(* IEC 61131-3 sources: StewartPlatform/Class/VaranManager (part 4) *)

    if (ud_LenObjName + ud_LenStr) < VARAN_MUTEX_NAME_MAX_LENGTH then
      _strcat(dest:=#str_CombinedName[0], src:=#str_ObjName[0]);
    else
      _strncpy(dest:=#str_ObjNamePart1[0], src:= #str_ObjName[0], max:= VARAN_MUTEX_NAME_MAX_LENGTH - ud_LenStr - ud_SepLenStr - VARAN_MUTEX_NAME_END_LENGTH - 1);    // Copy Beginning of str_ObjName
      _strncpy(dest:=#str_ObjNamePart2[0], src:= #str_ObjName[ud_LenObjName-VARAN_MUTEX_NAME_END_LENGTH-1], max:=VARAN_MUTEX_NAME_END_LENGTH);  // Copy Last MUTEX_NAME_END_LENGTH Char of str_ObjName

      // Put the Mutex String together
      _strcat(dest:=#str_CombinedName[0], src:= #str_ObjNamePart1[0]);
      _strcat(dest:=#str_CombinedName[0], src:= VARAN_STR_MUTEX_NAME_SEPERATOR);
      _strcat(dest:=#str_CombinedName[0], src:= #str_ObjNamePart2[0]);
    end_if;

    pv_RetMutex := OS_MT_CreateSemaphore(MTSEMATYPE_MUTEX, 1, 0, #str_CombinedName[0]);

    if pv_RetMutex = nil then

      // If Create Mutex failed: Insert the this pointer into the string
      ud_LenCombObjName := _strlen(#str_CombinedName[0]);

      str_this[0] := '%';
      str_this[1] := 'm';
      _itoa(udNumber:=pthis$UDINT, pString:=#str_this[2]);
      ud_LenThis  := _strlen(src:=#str_this[0]);

      _strcpy(dest:=#str_CombinedName[ud_LenCombObjName-ud_LenThis], src:=#str_this[0]);

      pv_RetMutex := OS_MT_CreateSemaphore(MTSEMATYPE_MUTEX, 1, 0, #str_CombinedName[0]);

    end_if;

  end_if;

END_FUNCTION

FUNCTION GLOBAL VaranManager::MutexStart
  VAR_INPUT
    pMutex 	: pVoid;
  END_VAR

  if(pMutex <> NIL) then
    OS_MT_WAIT(pMutex);
  end_if;

END_FUNCTION

FUNCTION GLOBAL VaranManager::MutexStop
  VAR_INPUT
    pMutex 	: pVoid;
  END_VAR

  if(pMutex <> NIL) then
    OS_MT_SIGNAL(pMutex);
  end_if;

END_FUNCTION
#endif

FUNCTION VIRTUAL GLOBAL VaranManager::Control::NewInst
  VAR_INPUT
    pPara 	: ^CmdStruct;
    pResult 	: ^Results;
  END_VAR
  VAR_OUTPUT
    ret_code 	: IprStates;
  END_VAR
  VAR
    p_paraAddDO           : ^t_VM_CMD_AddDO;
    p_paraMovDO           : ^t_VM_CMD_AddMovDo;
    p_paraGetPointers     : ^t_VM_CMD_GetDataPointers;
    p_paraGetModuleHandel : ^t_VM_CMD_GetModuleHandle;
    PostInitRetcode       : iprStates;
    pHelpPostInit         : ^t_s_PostInitList;
    i                     : UINT;

    pHelp                 : ^void;  // This pointer to call newinst
    // local variables for the Requested HWTString
    pStr_HWTRequested     : ^CHAR;
    ui_HWTRequestedLength : UINT;
    us_HWTRequestedCurrIndex  : USINT;
    i_Req                 :UINT;
    // local variables for HWTStrings in the VM
    pStr_HWTVM            : ^CHAR;
    us_HWTVMLength        : USINT;
    i_VM                  : USINT;
    ud_ModuleIndex        : UDINT;
    b_ModuleFound         : BOOL;

    // local variables to safe currently found module
    pStr_HWTVMCurrent     : ^CHAR;
    ud_ModuleIndexCurrent : UDINT;

    TempArray         : ARRAY [0..SERNO_STRING_SIZE-1] OF USINT;
    a_HelpArray       : ARRAY[0..99] OF CHAR;
	  ud_StrSize : UDINT;
    ud_MaxStrSize : UDINT;
    sSPIIDHeader  : t_s_SPIListHeader;

    //local variables for dummy mux callback
    sd_retval           :DINT;
  END_VAR

  ret_code := READY;  // Overwritten on error

  CASE pPara^.uiCmd OF
//**********************************************************************************************************************************************************
    CMD_POST_INIT_CALL: // call from hwcontrol
      // Check Loader Version if function is supported
      if ops.uiLoaderVersion$UINT >= VM_POST_INIT_AVAILABLE then
        bPostInitActive := TRUE;

#ifdef _LSL_TARGETARCH_ARM  // IO Image only needed for ARM  CPUs
#ifdef VARAN_iSetOutputImage
        // the image is not copied from the shadow ram to the VM DPRAM so far => copy it
        if (b_IOImageWritten = FALSE) & b_IOImage then
          VARAN_iSetOutputImage(VaranManagerNr, VARAN_DOL_ASY);
          b_IOImageWritten := TRUE;
        end_if;
#endif
#endif

        // we wait here until the initialisation of the Varan Rt and the SDIAS Clients has been finished
        CyWork(0);

        if bPostInitModulesReady then
          ret_code := READY;
          bPostInitActive := FALSE;
        else
          ret_code := BUSY;
        end_if;
      else
        // Should be impossible as we never request a Postinit if the Loader version is incorrect.
        TRACE("(VaranManager::Control::NewInst) CMD_POST_INIT_CALL not supported with current Loader. Loader Version >= 02.02.137 is required");
        ret_code := ERROR;
      end_if;

//**********************************************************************************************************************************************************
    CMD_POST_INIT_RT_SYNC:
      // check if all modules are ready
      if WaitForSyncSendObjectsCnt then
        CyWork(0);

        ret_code := BUSY;
      end_if;

//**********************************************************************************************************************************************************
    CMD_POST_INIT_RT_READY:
      // check post init modules
      if PostInitModuleCnt then
        pHelpPostInit := #aPostInitList[0];
        for i := 0 to PostInitModuleCnt - 1 do

          //call class, if it's still not ready
          if pHelpPostInit^.p_This then
            PostInitRetcode := pHelpPostInit^.p_This^.NewInst(pPara, pResult);

            // only overwrite the ready returncode if the returncode from the post init objects is different to it
            if PostInitRetcode <> READY then
              ret_code := PostInitRetcode;
            end_if;
          end_if;

          // set pointer on next this pointer
          pHelpPostInit += sizeof(t_s_PostInitList);
        end_for;
      end_if;

      // if manager is disabled => return error
      if ManagerOn = 0 then
        ret_code := ERROR;

      // if we're not ready, return busy
      elsif us_RtStep <> _RtWork then
        ret_code := BUSY;

      elsif ret_code = READY then
        // everything ready
        b_PostInitRtSyncReady := TRUE;
      end_if;

//**********************************************************************************************************************************************************
    CMD_FORCE_POST_INIT_END:  // call from hwcontrol
      // HWControl has run into timeout and has ended the Post Init Phase
      // This call informs the VM thats the Phase has ended.
      bPostInitActive := FALSE;

//**********************************************************************************************************************************************************
    CMD_POST_INIT_DO_SORT:    // call from hwcontrol
      // sort safety DOs if there is more than 1
      if pPriorityList & pPriorityList^.pNext &
        b_PayloadSupport = false then     // OS Handles Priorities of DO if b_PayloadSupport = true

        SortCmdsByPriority();

#ifdef _LSL_TARGETARCH_ARM  // IO Image only needed for ARM  CPUs
#ifdef VARAN_iSetOutputImage
        // Varandata has to be written once after sorting the DOs
        if b_IOImage then
          VARAN_iSetOutputImage(VaranManagerNr, VARAN_DOL_ISO);
        end_if;
      else
        // Varandata has to be written once after adding the DOs even without sorting anything because we need the shadow RAM image in the VM DPRAM)
        if b_IOImage then
          VARAN_iSetOutputImage(VaranManagerNr, VARAN_DOL_ISO);
        end_if;
#endif
#endif
      end_if;
//**********************************************************************************************************************************************************
    CMD_GET_HARDWARE_TREE_ENTRY:

      pHelp                 := nil;  // This pointer to call newinst
      // local variables for the Requested HWTString
      ui_HWTRequestedLength := 0;
      us_HWTRequestedCurrIndex  := 0;
      i_Req                 := 0;
      // local variables for HWTStrings in the VM
      pStr_HWTVM            := NIL;
      us_HWTVMLength        := 0;
      i_VM                  := 0;
      ud_ModuleIndex        := 0;
      b_ModuleFound         := FALSE;

      // local variables to safe currently found module
      pStr_HWTVMCurrent     := NIL;
      ud_ModuleIndexCurrent := 0;

      ret_code := ERROR;
      pResult^.aData[0]$t_HWCGetHardwareTreeEntryOut.retcode := _HWC_RETVAL_ERROR_VARAN_MODULE_NOT_FOUND;

      pStr_HWTRequested     := pPara^.aPara[0]$t_HWCGetHardwareDiagnosisIn.pStr_HardewareTreeEntry;

      //First HWT Path
      if pStr_HWTRequested = nil then

        ud_VaranPosition := VM_OBJECT_PATH;

        // Return String of the Varanmanger
        ret_code := READY;
        pResult^.aData$t_HWCGetHardwareTreeEntryOut.retcode := _HWC_RETVAL_OK_HWTSTR_RETURNED;
        pResult^.aData[0]$t_HWCGetHardwareTreeEntryOut.pStr_NextHardewareTreeEntry := (#ud_VaranPosition)$^CHAR;

      // Only possible for VM own HWT Path
      elsif (pStr_HWTRequested^$USINT = 2) then

        if pStr_HWTRequested^$UDINT = VM_OBJECT_PATH then

          if s_ModuleList.p_ModuleList^ then
            // Return first Module in list
            ret_code := s_ModuleList.p_ModuleList^$p_VaranBase^.NewInst(pPara,pResult);
          else
            // VM was found but there are no modules connected
            ret_code := READY;
            pResult^.aData[0]$t_HWCGetHardwareTreeEntryOut.retcode := _HWC_RETVAL_OK_MODULE_FOUND;
          end_if;
        end_if;

      else

        //Search for module
        ui_HWTRequestedLength     := (pStr_HWTRequested)$^UINT^ + 1;  //+1 because we compare the strings, 2 byte length
        us_HWTRequestedCurrIndex  := pPara^.aPara[0]$t_HWCGetHardwareDiagnosisIn.us_current_index;

        ud_ModuleIndex := 0;
        b_ModuleFound := FALSE;

        //loop over all modules
        while (ud_ModuleIndex < s_ModuleList.ud_NrOfModules) &
              (b_ModuleFound = FALSE) do

          pStr_HWTVM := (s_ModuleList.p_PositionList+ (ud_ModuleIndex * 4))^$^CHAR;  // 4 = SizeOf(^CHAR)

          if pStr_HWTVM  then
            us_HWTVMLength := pStr_HWTVM^;  //First byte is length

            i_Req := us_HWTRequestedCurrIndex;
            i_Vm  := 1;

            //Loop over strings
            while i_Req <= ui_HWTRequestedLength &
                  i_Vm  <= us_HWTVMLength do

              if (pStr_HWTRequested + i_Req)^ <> (pStr_HWTVM + i_Vm)^ then // Compare byte
                // Strings are not equal
                exit;
              end_if;

              i_Req += 1;
              i_VM  += 1;
            end_while;

            if (i_Req <= ui_HWTRequestedLength ) &                        // End of requested string was not reached
               (i_Vm = us_HWTVMLength + 1) &                              // And end of compared string reached
               ( (pStr_HWTRequested + i_Req)^ and HWT_ESCAPE_SEQU ) then  // Escape sequece found in Requested string

              b_ModuleFound := TRUE;

//              pPara^.aPara[0]$t_HWCGetHardwareDiagnosisIn.us_current_index   := i_Req$USINT;
//              pPara^.aPara[0]$t_HWCGetHardwareDiagnosisIn.us_current_length  := (ui_HWTRequestedLength - i_Req)$USINT;
              exit;
            end_if;

            if (i_Vm = us_HWTVMLength + 1) & (i_Req = ui_HWTRequestedLength + 1) then   // All Bytes and Length are equal
              b_ModuleFound := TRUE;
#ifdef HWK_SHOW_PRAGMA_MESSAGES
              #pragma message("LanSte 26.06.2014 16:11 \ check")
#endif

//              pPara^.aPara[0]$t_HWCGetHardwareDiagnosisIn.us_current_index  := i_Req$USINT - 1;  // -1 because we increased over max length at the end of the while loop
//              pPara^.aPara[0]$t_HWCGetHardwareDiagnosisIn.us_current_length := 1; // Last entry of string was reached, index points to last entry
              exit;
            end_if;

          end_if;

          ud_ModuleIndex += 1;  // Select next Module

        end_while;

        if b_ModuleFound then

          // Call module again incase it is an extension module
          pHelp := s_ModuleList.p_ModuleList + sizeof(p_VaranBase) * ud_ModuleIndex;
          ret_code := pHelp^$p_VaranBase^.NewInst(pPara,pResult);

          // Return if new HWT String was found
          if ret_code = READY &
             pResult^.aData[0]$t_HWCGetHardwareDiagnosisOut.retcode = _HWC_RETVAL_OK_HWTSTR_RETURNED then
            return;
          end_if;

          ud_ModuleIndex += 1;  // Select next Module
          ud_ModuleIndexCurrent := ud_ModuleIndex;

          b_ModuleFound := TRUE;  // Only set to enter loop

          while (ud_ModuleIndexCurrent < s_ModuleList.ud_NrOfModules) &
                (b_ModuleFound = TRUE) do

            pStr_HWTVMCurrent := (s_ModuleList.p_PositionList+ (ud_ModuleIndexCurrent * 4))^$^CHAR ;  // 4 = SizeOf(^CHAR)

            if pStr_HWTVMCurrent then

              // Check if module has already been called (multiple entries in list)
              ud_ModuleIndex := 0;
              b_ModuleFound := FALSE;

              //loop over all modules to search for duplicates
              while (ud_ModuleIndex < ud_ModuleIndexCurrent &
                     b_ModuleFound = FALSE) do

                pStr_HWTVM := (s_ModuleList.p_PositionList+ (ud_ModuleIndex * 4))^$^CHAR ;  // 4 = SizeOf(^CHAR)

                if pStr_HWTVM then

                  // Compare string length
                  if pStr_HWTVMCurrent^ = pStr_HWTVM^ then

                    // Compare string content
                    if _memcmp( ptr1 := pStr_HWTVMCurrent + 1,
                                ptr2 := pStr_HWTVM +1,
                                cntr := pStr_HWTVMCurrent^) = 0 then

                      // Multiple entry, Check next Module
                      b_ModuleFound := TRUE;
                      ud_ModuleIndexCurrent += 1;
                      exit;

                    end_if;
                  end_if;
                end_if;

                ud_ModuleIndex += 1;

              end_while;

              if b_ModuleFound = FALSE then
                exit; // Non duplicate entry
              end_if;

            else  // if pStr_HWTVMCurrent then
              ud_ModuleIndexCurrent += 1;
            end_if;

          end_while;

          if b_ModuleFound = FALSE then
            // Call Class
            pHelp := s_ModuleList.p_ModuleList + sizeof(p_VaranBase) * ud_ModuleIndexCurrent;
            ret_code := pHelp^$p_VaranBase^.NewInst(pPara,pResult);
          end_if;

        else
          pResult^.aData[0]$t_HWCGetHardwareDiagnosisOut.retcode := _HWC_RETVAL_ERROR_VARAN_MODULE_NOT_FOUND;
          ret_code := ERROR;
        end_if;

      end_if;

//**********************************************************************************************************************************************************
    CMD_GET_HARDWARE_DIAGNOSIS:

      pHelp                 := nil;  // This pointer to call newinst
      // local variables for the Requested HWTString
      ui_HWTRequestedLength := 0;
      us_HWTRequestedCurrIndex  := 0;
      i_Req                 := 0;
      // local variables for HWTStrings in the VM
      pStr_HWTVM            := NIL;
      us_HWTVMLength        := 0;
      i_VM                  := 0;
      ud_ModuleIndex        := 0;
      b_ModuleFound         := FALSE;

      ret_code := ERROR;
      pResult^.aData[0]$t_HWCGetHardwareDiagnosisOut.retcode := _HWC_RETVAL_ERROR;

      pStr_HWTRequested     := pPara^.aPara[0]$t_HWCGetHardwareDiagnosisIn.pStr_HardewareTreeEntry;

      if pStr_HWTRequested then

        // Check for VM String
        if (pStr_HWTRequested)$^UINT^ = 2 then

          if (pStr_HWTRequested)$^UDINT^ = VM_OBJECT_PATH then

            TempArray[0] := 0;

            if this <> p_this then
              //Reset statemachine
              eSPISSW := _GetVendorName;
              //Save This pointer
              p_this := this;

              // Reset Flags
              bDiagnosisDataAvailableFlags.HWVersion   := FALSE;
              bDiagnosisDataAvailableFlags.VendorName  := FALSE;
              bDiagnosisDataAvailableFlags.DeviceName  := FALSE;
              bDiagnosisDataAvailableFlags.OrderingNo  := FALSE;
              bDiagnosisDataAvailableFlags.LicenseNo   := FALSE;
              bDiagnosisDataAvailableFlags.SerialNo    := FALSE;
            end_if;

            case eSPISSW of
            	_GetVendorName:
                ret_code$DINT := GetSPIDataFromID(  p_us_position_info:=#TempArray[0]
                                                  , udListID:= VM_SPI_VENDOR_NAME_ID
                                                  , pData:= #a_VendorName[0]
                                                  , udRequDataLength:= sizeof(a_VendorName)
                                                  , pIDHeader:= #sSPIIDHeader
                                                  );

                if ret_code = READY then

                  // Null Termination ----------------------------------------
                  ud_StrSize    := sSPIIDHeader.ListLength;
                  ud_MaxStrSize := sizeof(a_VendorName);

                  pResult^.aData[0]$t_HWCGetHardwareDiagnosisOut.pStr_VendorName  := (#a_VendorName)$^CHAR; // Will be overwritten if this pointer is not equal

                  (pResult^.aData[0]$t_HWCGetHardwareDiagnosisOut.pStr_VendorName + ud_MaxStrSize)^ := 0;
                  if ud_StrSize < ud_MaxStrSize then
                    (pResult^.aData[0]$t_HWCGetHardwareDiagnosisOut.pStr_VendorName + ud_StrSize)^ := 0;
                  end_if;

                  bDiagnosisDataAvailableFlags.VendorName := TRUE;

                  eSPISSW := _GetSerialNo;
                  ret_code := BUSY;
                else
                  pResult^.aData[0]$t_HWCGetHardwareDiagnosisOut.retcode := _HWC_RETVAL_ERROR_VARAN_SPI_ACCESS_FAILED;
                  //set SSW to SPI Data Ready, because we return the values which are already in the HWK
                  eSPISSW := _SPIDataReady;
                  ret_code := BUSY;
                end_if;

              _GetSerialNo:
                ret_code$DINT := GetSPIDataFromID(  p_us_position_info:=#TempArray[0]
                                                  , udListID:= VM_SPI_SERIALNO_ID
                                                  , pData:= #a_SerialNo[0]
                                                  , udRequDataLength:= sizeof(a_SerialNo)
                                                  , pIDHeader:= #sSPIIDHeader
                                                  );

                if ret_code = READY then

                  // Null Termination ----------------------------------------
                  ud_StrSize    := sSPIIDHeader.ListLength;
                  ud_MaxStrSize := sizeof(a_SerialNo);

                  pResult^.aData[0]$t_HWCGetHardwareDiagnosisOut.pStr_SerialNo  := (#a_SerialNo)$^CHAR; // Will be overwritten if this pointer is not equal

                  (pResult^.aData[0]$t_HWCGetHardwareDiagnosisOut.pStr_SerialNo + ud_MaxStrSize)^ := 0;
                  if ud_StrSize < ud_MaxStrSize then
                    (pResult^.aData[0]$t_HWCGetHardwareDiagnosisOut.pStr_SerialNo + ud_StrSize)^ := 0;
                  end_if;

                  bDiagnosisDataAvailableFlags.SerialNo := TRUE;

                  eSPISSW := _GetDeviceName;
                  ret_code := BUSY;
                else
                  pResult^.aData[0]$t_HWCGetHardwareDiagnosisOut.retcode := _HWC_RETVAL_ERROR_VARAN_SPI_ACCESS_FAILED;
                  //set SSW to SPI Data Ready, because we return the values which are already in the HWK
                  eSPISSW := _SPIDataReady;
                  ret_code := BUSY;
                end_if;

            	_GetDeviceName:
                ret_code$DINT := GetSPIDataFromID(  p_us_position_info:=#TempArray[0]
                                                  , udListID:= VM_SPI_DEVICE_NAME_ID
                                                  , pData:= #a_DeviceName[0]
                                                  , udRequDataLength:= sizeof(a_DeviceName)
                                                  , pIDHeader:= #sSPIIDHeader
                                                  );

                if ret_code = READY then

                  // Null Termination ----------------------------------------
                  ud_StrSize    := sSPIIDHeader.ListLength;
                  ud_MaxStrSize := sizeof(a_DeviceName);

                  pResult^.aData[0]$t_HWCGetHardwareDiagnosisOut.pStr_DeviceName  := (#a_DeviceName)$^CHAR; // Will be overwritten if this pointer is not equal

                  (pResult^.aData[0]$t_HWCGetHardwareDiagnosisOut.pStr_DeviceName + ud_MaxStrSize)^ := 0;
                  if ud_StrSize < ud_MaxStrSize then
                    (pResult^.aData[0]$t_HWCGetHardwareDiagnosisOut.pStr_DeviceName + ud_StrSize)^ := 0;
                  end_if;

                  bDiagnosisDataAvailableFlags.DeviceName := TRUE;

                  eSPISSW := _GetOrderingNo;
                  ret_code := BUSY;
                else
                  pResult^.aData[0]$t_HWCGetHardwareDiagnosisOut.retcode := _HWC_RETVAL_ERROR_VARAN_SPI_ACCESS_FAILED;
                  //set SSW to SPI Data Ready, because we return the values which are already in the HWK
                  eSPISSW := _SPIDataReady;
                  ret_code := BUSY;
                end_if;

            	_GetOrderingNo:
                ret_code$DINT := GetSPIDataFromID(  p_us_position_info:=#TempArray[0]
                                                  , udListID:= VM_SPI_ORDERING_NO_ID
                                                  , pData:= #a_OrderingNo[0]
                                                  , udRequDataLength:= sizeof(a_OrderingNo)
                                                  , pIDHeader:= #sSPIIDHeader
                                                  );

                if ret_code = READY then

                  // Null Termination ----------------------------------------
                  ud_StrSize    := sSPIIDHeader.ListLength;
                  ud_MaxStrSize := sizeof(a_OrderingNo);

                  pResult^.aData[0]$t_HWCGetHardwareDiagnosisOut.pStr_OrderingNo  := (#a_OrderingNo)$^CHAR; // Will be overwritten if this pointer is not equal

                  (pResult^.aData[0]$t_HWCGetHardwareDiagnosisOut.pStr_OrderingNo + ud_MaxStrSize)^ := 0;
                  if ud_StrSize < ud_MaxStrSize then
                    (pResult^.aData[0]$t_HWCGetHardwareDiagnosisOut.pStr_OrderingNo + ud_StrSize)^ := 0;
                  end_if;

                  bDiagnosisDataAvailableFlags.OrderingNo := TRUE;

                  eSPISSW := _GetLicenseNoHWVersion;
                  ret_code := BUSY;
                else
                  pResult^.aData[0]$t_HWCGetHardwareDiagnosisOut.retcode := _HWC_RETVAL_ERROR_VARAN_SPI_ACCESS_FAILED;
                  //set SSW to SPI Data Ready, because we return the values which are already in the HWK
                  eSPISSW := _SPIDataReady;
                  ret_code := BUSY;
                end_if;

            	_GetLicenseNoHWVersion:

                ret_code$DINT := GetSPIDataFromID(  p_us_position_info:=#TempArray[0]
                                                  , udListID:= VM_SPI_IDENTIFICATION_LIST
                                                  , pData:= #a_HelpArray[0]
                                                  , udRequDataLength:= sizeof(udHWVersion) + sizeof(udLicenseNo)
                                                  , pIDHeader:= #sSPIIDHeader
                                                  , udOffset := 8
                                                  );

                udLicenseNo := a_HelpArray[0]$UDINT;
                udHWVersion := a_HelpArray[4]$UDINT;

                if ret_code = READY then
                  bDiagnosisDataAvailableFlags.LicenseNo := TRUE;
                  bDiagnosisDataAvailableFlags.HWVersion := TRUE;
                  eSPISSW := _SPIDataReady;
                  ret_code := BUSY;
                else
                  pResult^.aData[0]$t_HWCGetHardwareDiagnosisOut.retcode := _HWC_RETVAL_ERROR_VARAN_SPI_ACCESS_FAILED;
                  //set SSW to SPI Data Ready, because we return the values which are already in the HWK
                  eSPISSW := _SPIDataReady;
                  ret_code := BUSY;
                end_if;

            	_SPIDataReady:
                //Don't reset statemachine because if we have the same this pointer we don't have to make spi Accesses again
                //eSPISSW := _GetVendorName;

                //Data which is already in HWK available
                if p_NodeInfo then

                  pResult^.aData$t_HWCGetHardwareDiagnosisOut.hd_FPGAVersion  := to_udint(p_NodeInfo^.ucFPGAVersion);
                  pResult^.aData$t_HWCGetHardwareDiagnosisOut.ud_DeviceID     := to_udint(p_NodeInfo^.uiDeviceID);
                  pResult^.aData$t_HWCGetHardwareDiagnosisOut.ud_VendorID     := to_udint(p_NodeInfo^.uiVendorID);
                end_if;

                if bDiagnosisDataAvailableFlags.VendorName then
                  pResult^.aData[0]$t_HWCGetHardwareDiagnosisOut.pStr_VendorName  := (#a_VendorName)$^CHAR;
                end_if;

                if bDiagnosisDataAvailableFlags.HWVersion & bDiagnosisDataAvailableFlags.LicenseNo then
                  pResult^.aData[0]$t_HWCGetHardwareDiagnosisOut.hd_HWVersion     := udHWVersion;
                  pResult^.aData[0]$t_HWCGetHardwareDiagnosisOut.ud_LicenseNo      := udLicenseNo;
                end_if;

                if bDiagnosisDataAvailableFlags.DeviceName then
                  pResult^.aData[0]$t_HWCGetHardwareDiagnosisOut.pStr_DeviceName  := (#a_DeviceName)$^CHAR;
                end_if;

                if bDiagnosisDataAvailableFlags.OrderingNo then
                  pResult^.aData[0]$t_HWCGetHardwareDiagnosisOut.pStr_OrderingNo  := (#a_OrderingNo)$^CHAR;
                end_if;

                if bDiagnosisDataAvailableFlags.SerialNo then
                  pResult^.aData[0]$t_HWCGetHardwareDiagnosisOut.pStr_SerialNo := (#a_SerialNo)$^CHAR;
                end_if;

                ret_code := READY;
                pResult^.aData[0]$t_HWCGetHardwareDiagnosisOut.retcode := _HWC_RETVAL_OK;

            end_case;
          end_if;

          return;
        end_if;

        ui_HWTRequestedLength     := (pStr_HWTRequested)$^UINT^ + 1;  //+1 because we compare the strings, 2 byte length
        us_HWTRequestedCurrIndex  := pPara^.aPara[0]$t_HWCGetHardwareDiagnosisIn.us_current_index;

        ud_ModuleIndex := 0;
        b_ModuleFound := FALSE;

        //loop over all modules
        while (ud_ModuleIndex < s_ModuleList.ud_NrOfModules) &
              (b_ModuleFound = FALSE) do

          pStr_HWTVM := (s_ModuleList.p_PositionList+ (ud_ModuleIndex * 4))^$^CHAR ;  // 4 = SizeOf(^CHAR)

          if pStr_HWTVM  then
            us_HWTVMLength := pStr_HWTVM^;  //First byte is length

            i_Req := us_HWTRequestedCurrIndex;
            i_Vm  := 1;

            //Loop over strings
            while i_Req <= ui_HWTRequestedLength &
                  i_Vm  <= us_HWTVMLength do

//              if (pStr_HWTRequested + i_Req)^ and HWT_ESCAPE_SEQU then  // Check for Escape Sequenze
//                b_ModuleFound := TRUE;
//                exit;
//              end_if;

              if (pStr_HWTRequested + i_Req)^ <> (pStr_HWTVM + i_Vm)^ then // Compare byte
                // Strings are not equal
                exit;
              end_if;

              i_Req += 1;
              i_VM  += 1;
            end_while;

//            #pragma message("LanSte 18.06.2014 18:23 \ Index Update testen")
//            if b_ModuleFound then // Escape Sequence was found
//
//              pPara^.aPara[0]$t_HWCGetHardwareDiagnosisIn.us_current_index   := i_Req$USINT;
//              pPara^.aPara[0]$t_HWCGetHardwareDiagnosisIn.us_current_length  := (ui_HWTRequestedLength - i_Req)$USINT;
//              exit;
//
//            end_if;

            if (i_Req <= ui_HWTRequestedLength ) &                        // End of requested string was not reached
            (i_Vm = us_HWTVMLength + 1) &                                 // And end of compared string reached
               ( (pStr_HWTRequested + i_Req)^ and HWT_ESCAPE_SEQU ) then  // Escape sequece found in Requested string

              b_ModuleFound := TRUE;
              pPara^.aPara[0]$t_HWCGetHardwareDiagnosisIn.us_current_index   := i_Req$USINT;
              pPara^.aPara[0]$t_HWCGetHardwareDiagnosisIn.us_current_length  := (ui_HWTRequestedLength - i_Req)$USINT;
              exit;
            end_if;

            if (i_Vm = us_HWTVMLength + 1) & (i_Req = ui_HWTRequestedLength + 1) then   // All Bytes and Length are equal
              b_ModuleFound := TRUE;
              pPara^.aPara[0]$t_HWCGetHardwareDiagnosisIn.us_current_index  := i_Req$USINT - 1;  // -1 because we increased over max length at the end of the while loop
              pPara^.aPara[0]$t_HWCGetHardwareDiagnosisIn.us_current_length := 1; // Last entry of string was reached, index points to last entry
              exit;
            end_if;

          end_if;

          ud_ModuleIndex += 1;  // Select next Module

        end_while;

        if b_ModuleFound then
          // Call Class
          pHelp := s_ModuleList.p_ModuleList + sizeof(p_VaranBase) * ud_ModuleIndex;
          ret_code := pHelp^$p_VaranBase^.NewInst(pPara,pResult);
        else
          pResult^.aData[0]$t_HWCGetHardwareDiagnosisOut.retcode := _HWC_RETVAL_ERROR_VARAN_MODULE_NOT_FOUND;
          ret_code := ERROR;
        end_if;

      end_if;

//**********************************************************************************************************************************************************
    VM_CMD_NEED_POST_INIT_CALL: // call from varan client
      // Check Loader Version if function is supported
      if ops.uiLoaderVersion$UINT >= VM_POST_INIT_AVAILABLE then

        // store this pointer of the module
        aPostInitList[PostInitModuleCnt].p_This := pPara^.aPara[0]$p_VaranBase;

        // remember if we have to wait for DOs to be created
        aPostInitList[PostInitModuleCnt].Settings := pPara^.aPara[1]$BSINT;
        if aPostInitList[PostInitModuleCnt].Settings.Wait4DOCreation then
          WaitForPostInitObjectsCnt += 1;
          if aPostInitList[PostInitModuleCnt].Settings.Wait4MoveDOCreation then
            WaitForPostInitMoveObjectsCnt += 1;
          end_if;
        end_if;

        // remember if we have to wait for the sync of this module
        if aPostInitList[PostInitModuleCnt].Settings.Wait4SyncSend then
          WaitForSyncSendObjectsCnt += 1;
        end_if;

        aPostInitList[PostInitModuleCnt].b_CallMe := TRUE;

        // return index for this module
        pResult^.uiLng := 2;
        pResult^.aData[0]$UINT := PostInitModuleCnt;

        // increase number of post init modules
        PostInitModuleCnt += 1;

        // we're no longer ready with post init. we have to wait until all modules from the list are finished
        bPostInitModulesReady := FALSE;
      else
        TRACE("(VaranManager::Control::NewInst) VM_CMD_NEED_POST_INIT_CALL not supported with current Loader. Loader Version >= 02.02.137 is required");
        ret_code := ERROR;
      end_if;

//**********************************************************************************************************************************************************
    VM_CMD_POST_INIT_FINISHED: // call from varan client
      // Check Loader Version if function is supported
      if ops.uiLoaderVersion$UINT >= VM_POST_INIT_AVAILABLE then

        // only relevant during last Init
        if PostInitModuleCnt then
          // check if it's a valid index
          if pPara^.aPara[1]$UINT < VM_MAX_POST_INIT_MODULES then
            // check if our local this pointer matches this object
            if pPara^.aPara[0]$p_VaranBase = aPostInitList[pPara^.aPara[1]$UINT].p_This then
              // increase number of ready objects
              PostInitModuleReadyCnt += 1;
//              aPostInitList[pPara^.aPara[1]$UINT].b_CallMe := FALSE;

              // check if it's an object we were waiting for
              if aPostInitList[pPara^.aPara[1]$UINT].Settings.Wait4DOCreation then
                aPostInitList[pPara^.aPara[1]$UINT].Settings.Wait4DOCreation := FALSE;

                if WaitForPostInitObjectsCnt then
                  WaitForPostInitObjectsCnt -= 1;
                else
                  TRACE("(VaranManager::Control::NewInst) There is already no more post init object to wait for! (VM_CMD_POST_INIT_FINISHED)");
                  ret_code := ERROR;
                end_if;
              end_if;

              // check if it's an object we were waiting for
              if aPostInitList[pPara^.aPara[1]$UINT].Settings.Wait4MoveDOCreation then
                aPostInitList[pPara^.aPara[1]$UINT].Settings.Wait4MoveDOCreation := FALSE;

                if WaitForPostInitMoveObjectsCnt then
                  WaitForPostInitMoveObjectsCnt -= 1;
                else
                  TRACE("(VaranManager::Control::NewInst) There is already no more post init object to wait for (create move DOs)! (VM_CMD_POST_INIT_FINISHED)");
                  ret_code := ERROR;
                end_if;
              end_if;

              // on last init we check if all modules which need to have finished their init
              if PostInitModuleReadyCnt = PostInitModuleCnt then
                bPostInitModulesReady := TRUE;
              end_if;
            else
              TRACE("(VaranManager::Control::NewInst) This pointer of post init module given doesn't match locally stored this pointer for this index!");
              ret_code := ERROR;
            end_if;
          else
            TRACE("(VaranManager::Control::NewInst) Invalid index of post init module given!");
            ret_code := ERROR;
          end_if;
        else
          TRACE("(VaranManager::Control::NewInst) More modules ready with last init than expected");
          ret_code := ERROR;
        end_if;
      else
        TRACE("(VaranManager::Control::NewInst) VM_CMD_POST_INIT_FINISHED not supported with current Loader. Loader Version >= 02.02.137 is required");
        ret_code := ERROR;
      end_if;

//**********************************************************************************************************************************************************
    VM_CMD_IS_PAYLOAD_SUPPORTED:  // to get the status of PayloadSupport
      pResult^.aData[0]$BOOL := b_PayloadSupport;

//**********************************************************************************************************************************************************
    VM_CMD_DO_CREATION_FINISHED: // a post-init module is finished with creating DOs
      // Check Loader Version if function is supported
      if ops.uiLoaderVersion$UINT >= VM_POST_INIT_AVAILABLE then

        // only relevant during last Init
        if PostInitModuleCnt then
          // check if it's a valid index
          if pPara^.aPara[1]$UINT < VM_MAX_POST_INIT_MODULES then
            // check if our local this pointer matches this object
            if pPara^.aPara[0]$p_VaranBase = aPostInitList[pPara^.aPara[1]$UINT].p_This then
              // check if it's an object we were waiting for
              if aPostInitList[pPara^.aPara[1]$UINT].Settings.Wait4DOCreation then
                aPostInitList[pPara^.aPara[1]$UINT].Settings.Wait4DOCreation := FALSE;

                if WaitForPostInitObjectsCnt then
                  WaitForPostInitObjectsCnt -= 1;
                else
                  TRACE("(VaranManager::Control::NewInst) There is already no more post init object to wait for!");
                  ret_code := ERROR;
                end_if;
              else
                TRACE("(VaranManager::Control::NewInst) Module finished with DO creation, where  There is already no more post init object to wait for!");
                ret_code := ERROR;
              end_if;
            else
              TRACE("(VaranManager::Control::NewInst) This pointer of post init module given doesn't match locally stored this pointer for this index!");
              ret_code := ERROR;
            end_if;
          else
            TRACE("(VaranManager::Control::NewInst) Invalid index of post init module given!");
            ret_code := ERROR;
          end_if;
        else
          TRACE("(VaranManager::Control::NewInst) More modules ready with last init than expected");
          ret_code := ERROR;
        end_if;
      else
        TRACE("(VaranManager::Control::NewInst) VM_CMD_DO_CREATION_FINISHED not supported with current Loader. Loader Version >= 02.02.137 is required");
        ret_code := ERROR;
      end_if;

//**********************************************************************************************************************************************************
    VM_CMD_MOVE_DO_CREATION_FINISHED:
      // Check Loader Version if function is supported
      if ops.uiLoaderVersion$UINT >= VM_POST_INIT_AVAILABLE then

        // only relevant during last Init
        if PostInitModuleCnt then
          // check if it's a valid index
          if pPara^.aPara[1]$UINT < VM_MAX_POST_INIT_MODULES then
            // check if our local this pointer matches this object
            if pPara^.aPara[0]$p_VaranBase = aPostInitList[pPara^.aPara[1]$UINT].p_This then
              // check if it's an object we were waiting for
              if aPostInitList[pPara^.aPara[1]$UINT].Settings.Wait4MoveDOCreation then
                aPostInitList[pPara^.aPara[1]$UINT].Settings.Wait4MoveDOCreation := FALSE;

                if WaitForPostInitMoveObjectsCnt then
                  WaitForPostInitMoveObjectsCnt -= 1;
                else
                  TRACE("(VaranManager::Control::NewInst) There is already no more post init object to wait for (create move DOs)!");
                  ret_code := ERROR;
                end_if;
              else
                TRACE("(VaranManager::Control::NewInst) Module finished with move DO creation, where  There is already no more post init object to wait for!");
                ret_code := ERROR;
              end_if;
            else
              TRACE("(VaranManager::Control::NewInst) This pointer of post init module given doesn't match locally stored this pointer for this index! (Move DOs)");
              ret_code := ERROR;
            end_if;
          else
            TRACE("(VaranManager::Control::NewInst) Invalid index of post init module given! (Move DOs)");
            ret_code := ERROR;
          end_if;
        else
          TRACE("(VaranManager::Control::NewInst) More modules ready with last init than expected (Move DOs)");
          ret_code := ERROR;
        end_if;
      else
        TRACE("(VaranManager::Control::NewInst) VM_CMD_MOVE_DO_CREATION_FINISHED not supported with current Loader. Loader Version >= 02.02.137 is required (Move DOs)");
        ret_code := ERROR;
      end_if;

//**********************************************************************************************************************************************************
    VM_CMD_DO_MEM_READY: // check if all post init objects are finished with creating DOs
      // if we're not in post init or the varan manager has finished waiting for post init objects => the DO memory is ready
      if WaitForPostInitObjectsCnt = 0 then
        pResult^.aData[4] := TRUE;
      else
        pResult^.aData[4] := FALSE;
      end_if;

//**********************************************************************************************************************************************************
    VM_CMD_MOVE_DO_MEM_READY: // check if all post init objects are finished with creating move DOs
      // if we're not in post init or the varan manager has finished waiting for post init objects => the move DO memory is ready
      if WaitForPostInitMoveObjectsCnt = 0 then
        pResult^.aData[4] := TRUE;
      else
        pResult^.aData[4] := FALSE;
      end_if;

//**********************************************************************************************************************************************************
    VM_CMD_SYNC_SEND_READY:
      // only work on it if the post init rt hasn't been finished, otherwise we would have the log messages if modules are plugged at runtime
      if b_PostInitRtSyncReady = FALSE then
        // Check Loader Version if function is supported
        if ops.uiLoaderVersion$UINT >= VM_POST_INIT_AVAILABLE then
          // only relevant during last Init
          if PostInitModuleCnt then
            // check if it's a valid index
            if pPara^.aPara[1]$UINT < VM_MAX_POST_INIT_MODULES then
              // check if our local this pointer matches this object
              if pPara^.aPara[0]$p_VaranBase = aPostInitList[pPara^.aPara[1]$UINT].p_This then
                // check if it's an object we were waiting for
                if aPostInitList[pPara^.aPara[1]$UINT].Settings.Wait4SyncSend then
                  aPostInitList[pPara^.aPara[1]$UINT].Settings.Wait4SyncSend := FALSE;

                  if WaitForSyncSendObjectsCnt then
                    WaitForSyncSendObjectsCnt -= 1;
                  else
                    TRACE("(VaranManager::Control::NewInst) There is already no more post init object to wait for (sync send ready)!");
                    ret_code := ERROR;
                  end_if;
                else
                  TRACE("(VaranManager::Control::NewInst) Module finished with sync send ready, where  There is already no more post init object to wait for!");
                  ret_code := ERROR;
                end_if;
              else
                TRACE("(VaranManager::Control::NewInst) This pointer of post init module given doesn't match locally stored this pointer for this index! (Move DOs)");
                ret_code := ERROR;
              end_if;
            else
              TRACE("(VaranManager::Control::NewInst) Invalid index of post init module given! (sync send ready)");
              ret_code := ERROR;
            end_if;
          else
            TRACE("(VaranManager::Control::NewInst) More modules ready with last init than expected (sync send ready)");
            ret_code := ERROR;
          end_if;
        else
          TRACE("(VaranManager::Control::NewInst) VM_CMD_MOVE_DO_CREATION_FINISHED not supported with current Loader. Loader Version >= 02.02.137 is required (Move DOs)");
          ret_code := ERROR;
        end_if;
      end_if;

//**********************************************************************************************************************************************************
    VM_CMD_SET_MUX_THIS: // ignore this command, it's only for the VaranMux classes
      ret_code := ERROR; // return error => command not handled

//**********************************************************************************************************************************************************
    VM_CMD_INSTALL_DUMMY_CALLBACK:

      if pPara^.aPara[0] >= 4 * sizeof(DINT) then

        sd_retval := AddObjectCallback(p_us_position_info:=pPara^.aPara[1]$^USINT
                        , ud_action_ptr:= pPara^.aPara[2]$UDINT
                        , ud_thisp:= pPara^.aPara[3]$UDINT
                        , sd_required:= pPara^.aPara[4]);
      else

        TRACE("(VaranManager::Control::NewInst) VM_CMD_INSTALL_DUMMY_CALLBACK. Length of NewInst Commando is invalid");
      end_if;

//**********************************************************************************************************************************************************
    else    // Commands for Payload
      if b_PayloadSupport then

        pResult^.uiLng := sizeof(DINT);
        pResult^.aData[0]$DINT := VM_CMD_NOT_IMPLEMENTED; // Default Return code, must be overwritten by induvidual methods

        CASE pPara^.uiCmd OF

        //*****************************************************************************
          VM_CMD_GET_MODULE_HANDLE :
            p_paraGetModuleHandel := (pPara^.aPara[0])$^t_VM_CMD_GetModuleHandle;

            pResult^.aData[0]$DINT := GetModuleHandle(  p_us_PositionInfo := p_paraGetModuleHandel^.p_us_position_info
                                                      , p_ud_ModuleHandle := p_paraGetModuleHandel^.p_ud_module_handle);

        //*****************************************************************************
          VM_CMD_ADD_DO :
            p_paraAddDO := (pPara^.aPara[0])$^t_VM_CMD_AddDO;
            pResult^.aData[0]$DINT := AddPayloadDO( p_ud_DoHandle                 := p_paraAddDO^.p_ud_DoHandle
                                                  , ud_NodeHandle                 := p_paraAddDO^.ud_ModuleHandle
                                                  , ud_DoRequired                 := p_paraAddDO^.ud_b_DoRequired
                                                  , ud_DolType                    := p_paraAddDO^.ud_DolType
                                                  , ud_Command                    := p_paraAddDO^.ud_Command
                                                  , ud_Priority                   := p_paraAddDO^.ud_Priority
                                                  , ud_PrescalerCounterThreshold  := p_paraAddDO^.ud_PreScalerCounterThreshold
                                                  , ud_PrescalerCounterStartValue := p_paraAddDO^.ud_PreScalerCounterStartValue
                                                  , ud_ReadOffset                 := p_paraAddDO^.ud_OffsetRead
                                                  , ud_ReadLength                 := p_paraAddDO^.ud_LengthRead
                                                  , ud_WriteOffset                := p_paraAddDO^.ud_OffsetWrite
                                                  , ud_WriteLength                := p_paraAddDO^.ud_LengthWrite
                                                  , ud_Filter                     := p_paraAddDO^.ud_Filter
                                                  , ud_Slices                     := p_paraAddDO^.ud_Slices
                                                  , ud_WritePayloadType           := p_paraAddDO^.ud_WritePayloadType);

        //*****************************************************************************
          VM_CMD_ADD_MOV_DO :
            p_paraMovDO := (pPara^.aPara[0])$^t_VM_CMD_AddMovDo;
            pResult^.aData[0]$DINT := AddPayloadMoveDO( p_ud_DoHandle                 := p_paraMovDO^.p_ud_DoHandle
                                                      , ud_bDoRequired                := p_paraMovDO^.ud_b_DoRequired
                                                      , ud_DolType                    := p_paraMovDO^.ud_DolType
                                                      , ud_Priority                   := p_paraMovDO^.ud_Priority
                                                      , ud_PrescalerCounterThreshold  := p_paraMovDO^.ud_PreScalerCounterThreshold
                                                      , ud_PrescalerCounterStartValue := p_paraMovDO^.ud_PreScalerCounterStartValue
                                                      , ud_hSourceReadDoHandle        := p_paraMovDO^.ud_SourceReadDoHandle
                                                      , ud_ReadOffset                 := p_paraMovDO^.ud_SourceReadOffset
                                                      , ud_hDestinationWriteDoHandle  := p_paraMovDO^.ud_DestinationWriteDoHandle
                                                      , ud_WriteOffset                := p_paraMovDO^.ud_DestinationWriteOffset
                                                      , ud_MoveDataLength             := p_paraMovDO^.ud_LengthMove);

        //*****************************************************************************
          VM_CMD_GET_DATA_POINTERS  :
            p_paraGetPointers := (pPara^.aPara[0])$^t_VM_CMD_GetDataPointers;
            pResult^.aData[0]$DINT := GetDataPointers(  ud_hDoHandle  := p_paraGetPointers^.ud_DoHandle
                                                      , pp_ReadData   := p_paraGetPointers^.p_ud_ReadData$^pVoid
                                                      , pp_WriteData  := p_paraGetPointers^.p_ud_WriteData$^pVoid);

        //*****************************************************************************
          VM_CMD_IS_DMA_ACTIVE :
            if PayloadFrame then
              pResult^.aData[0]$BOOL := TRUE;
            else
              pResult^.aData[0]$BOOL := FALSE;
            end_if;

          else
            ret_code := ERROR;
        END_CASE;

      else
        pResult^.uiLng := sizeof(DINT);
        pResult^.aData[0]$DINT := VM_CMD_NOT_IMPLEMENTED;
        TRACE("(VaranManager::Control::NewInst) Unknown command!");
        ret_code := ERROR;
      end_if;

  END_CASE;

END_FUNCTION

FUNCTION VaranManager::TurnOffIsoTask
  VAR
    s_PropertyValuePair : LSL_PROPERTY_VALUE_PAIR;
  END_VAR

  if b_PayloadSupport &
     _RTOSVersion >= VM_FULL_PAYLOAD_AVAILABLE  then
    s_PropertyValuePair.udPropertyId    := VM_PROP_TASK_STATE_ISO;
    s_PropertyValuePair.udPropertyValue := TK_STATE_STOPPED;
    MULTI_VARAN_iSetNodeProperties( hNodeHandle           := vmNodeHandle
                                  , udPropertyCount       := 1
                                  , psPropertyValuePairs  := #s_PropertyValuePair);
  else
    p_ManagerStructure^.ucTCEnable := p_ManagerStructure^.ucTCEnable AND VM_DISABLE_ISO_TASK;
  end_if;

END_FUNCTION

FUNCTION VaranManager::AddPayloadDO
  VAR_INPUT
    p_ud_DoHandle 	: ^UDINT;
    ud_NodeHandle 	: UDINT;
    ud_DoRequired 	: UDINT;
    ud_DolType 	: UDINT;
    ud_Command 	: UDINT;
    ud_Priority 	: UDINT;
    ud_PrescalerCounterThreshold 	: UDINT;
    ud_PrescalerCounterStartValue 	: UDINT;
    ud_ReadOffset 	: UDINT;
    ud_ReadLength 	: UDINT;
    ud_WriteOffset 	: UDINT;
    ud_WriteLength 	: UDINT;
    ud_Filter 	: UDINT;
    ud_Slices 	: UDINT;
    ud_WritePayloadType :  UDINT;
  END_VAR
  VAR_OUTPUT
    sd_retval 	: DINT;
  END_VAR
  VAR
    TempMem             :  UDINT;
    TempMemWr           :  UDINT;
  END_VAR

#ifdef VM_DEBUG_PAYLOAD
  if b_PayloadSupport = false then
    // This method is not suppored without payload
    ((0)$^USINT)^ := 0;
  end_if;
#endif

  //look if we Manager is on
  if ( ManagerOn ) then
    //look if we must execute Cyclic DOL list
    if ( ud_DolType = VARAN_DOL_ASY ) then
      s_CyHandles.b_ExecuteDOL := TRUE;			//set flag to execut Dol list
    end_if;

    sd_retval := MULTI_VARAN_iAddDo(  phDoHandle    := p_ud_DoHandle
                                    , hNodeHandle   := ud_NodeHandle
                                    , bDoRequired   := ud_DoRequired
                                    , udDolType     := ud_DolType
                                    , udCommand     := ud_Command
                                    , udPriority    := ud_Priority
                                    , udPrescalerCounterThreshold   := ud_PrescalerCounterThreshold
                                    , udPrescalerCounterStartValue  := ud_PrescalerCounterStartValue
                                    , udReadOffset  := ud_ReadOffset
                                    , udReadLength  := ud_ReadLength
                                    , udWriteOffset := ud_WriteOffset
                                    , udWriteLength := ud_WriteLength
                                    , udFilter      := ud_Filter
                                    , udSlices      := ud_Slices
                                    , udWritePayloadType := ud_WritePayloadType$LSL_WRITE_PAYLOAD_TYPE);

    //look if an error occured
    if ( sd_retval <> VARANMANAGER_OK ) then
      s_ErrorVaranManager.f_AddRdDO := SetVaranDOError( sd_Error 		:= sd_retval
                                                      , b_manager_off	:= TRUE
                                                      , b_log			:= TRUE
                                                      );
    else

      if PayloadFrame then  // Use PayloadFrame because, b_PayloadSupport only shows the interface used.
                            // Payload DO Mem Calculaition +++++++++++++++++++++++++++++++++++++++++++++++++++++++++++++++++++++++++++++++++++++++++++++++++++++++++++++++++++++++++++++++++++++++++
        case ud_Command of

            VARAN_CMD_CONTROL_READ,
            VARAN_CMD_MEMORY_READ:      // Read DO -------------------------------------------------------------------------------------------------------------------------------
                // 1 Byte Status + n Byte (Load data read) + 0 to 3 Byte (compensate missalignment)
                TempMem := 1 + ud_ReadLength;

                // 1 Byte Control
                TempMemWr := 1;

                // Increase for variable DO
                if ud_WritePayloadType > WR_PLD_TYPE_STANDARD$UDINT then
                  TempMemWr += 16#0D;
                end_if;

                case ud_DolType of
                // **************************************************
                  VARAN_DOL_DA:
                    DPRAM_Used.DA_Rd          += TempMem + TempMemWr + SIZE_PAYLOAD_FRAME_HEADER_DO;
                    DPRAM_Used_Payload.DA_Rd  += TempMem;
                    DPRAM_Used_Payload.DA_Wr  += TempMemWr;
                    DOCounter.DA_Rd  += 1;

                // **************************************************
                  VARAN_DOL_ISO:
                    DPRAM_Used.ISO_Rd         += TempMem + TempMemWr + SIZE_PAYLOAD_FRAME_HEADER_DO;
                    DPRAM_Used_Payload.ISO_Rd += TempMem;
                    DPRAM_Used_Payload.ISO_Wr += TempMemWr;
                    DOCounter.ISO_Rd  += 1;

                // **************************************************
                  VARAN_DOL_ASY:
                    DPRAM_Used.ASY_Rd         += TempMem + TempMemWr + SIZE_PAYLOAD_FRAME_HEADER_DO;
                    DPRAM_Used_Payload.ASY_Rd += TempMem;
                    DPRAM_Used_Payload.ASY_Wr += TempMemWr;
                    DOCounter.ASY_Rd  += 1;

                // **************************************************
                  VARAN_DOL_ADMIN:
                    DPRAM_Used.Admin_Rd         += TempMem + TempMemWr + SIZE_PAYLOAD_FRAME_HEADER_DO;
                    DPRAM_Used_Payload.Admin_Rd += TempMem;
                    DPRAM_Used_Payload.ASY_Wr   += TempMemWr;
                    DOCounter.Admin_Rd += 1;

                // **************************************************
                  VARAN_DOL_IRQ:
                    DPRAM_Used.IRQ_Rd         += TempMem + TempMemWr + SIZE_PAYLOAD_IRQ_FRAME_HEADER_DO;
                    DPRAM_Used_Payload.IRQ_Rd += TempMem;
                    DPRAM_Used_Payload.IRQ_Wr += TempMemWr;
                    DOCounter.IRQ_Rd  += 1;
                end_case;

                DPRAM_Used_Payload.Payload_Read += TempMem;
                DPRAM_Used_Payload.Payload_Write += TempMemWr;

                if ud_DolType <> VARAN_DOL_IRQ then
                  DPRAM_Used.Total  += TempMem + TempMemWr + SIZE_PAYLOAD_FRAME_HEADER_DO;
                  DPRAM_Used_Payload.Payload_Header += SIZE_PAYLOAD_FRAME_HEADER_DO;
                else
                  DPRAM_Used.Total  += TempMem + TempMemWr + SIZE_PAYLOAD_IRQ_FRAME_HEADER_DO;
                  DPRAM_Used_Payload.Payload_Header += SIZE_PAYLOAD_IRQ_FRAME_HEADER_DO;
                end_if;

                DPRAM_Used_Payload.Total  += TempMem + TempMemWr;

                DOCounter.Total   += 1;

            VARAN_CMD_CONTROL_WRITE,
            VARAN_CMD_MEMORY_WRITE:     // Write DO -------------------------------------------------------------------------------------------------------------------------------
                // 1 Byte Control + n Byte (Load data read) + 0 to 3 Byte (compensate missalignment)
                TempMemWr := 1 + ud_WriteLength;

                // Increase for variable DO
                if ud_WritePayloadType > WR_PLD_TYPE_STANDARD$UDINT then
                  TempMemWr += 16#0D;
                end_if;

                // 1 Byte Status in Read DPRAM
                TempMem := 1;

                case ud_DolType of
                // **************************************************
                  VARAN_DOL_DA:
                    DPRAM_Used.DA_Wr            += TempMem + TempMemWr + SIZE_PAYLOAD_FRAME_HEADER_DO;
                    DPRAM_Used_Payload.DA_Rd    += TempMem;
                    DPRAM_Used_Payload.DA_Wr    += TempMemWr;
                    DOCounter.DA_Wr  += 1;

                // **************************************************
                  VARAN_DOL_ISO:
                    DPRAM_Used.ISO_Wr           += TempMem + TempMemWr + SIZE_PAYLOAD_FRAME_HEADER_DO;
                    DPRAM_Used_Payload.ISO_Rd   += TempMem;
                    DPRAM_Used_Payload.ISO_Wr   += TempMemWr;
                    DOCounter.ISO_Wr += 1;

                // **************************************************
                  VARAN_DOL_ASY:
                    DPRAM_Used.ASY_Wr           += TempMem + TempMemWr + SIZE_PAYLOAD_FRAME_HEADER_DO;
                    DPRAM_Used_Payload.ASY_Rd   += TempMem;
                    DPRAM_Used_Payload.ASY_Wr   += TempMemWr;
                    DOCounter.ASY_Wr  += 1;

                // **************************************************
                  VARAN_DOL_ADMIN:
                    DPRAM_Used.Admin_Wr         += TempMem + TempMemWr + SIZE_PAYLOAD_FRAME_HEADER_DO;
                    DPRAM_Used_Payload.Admin_Rd += TempMem;
                    DPRAM_Used_Payload.Admin_Wr += TempMemWr;
                    DOCounter.Admin_Wr  += 1;

                // **************************************************
                  VARAN_DOL_IRQ:
                    DPRAM_Used.IRQ_Wr           += TempMem + TempMemWr + SIZE_PAYLOAD_IRQ_FRAME_HEADER_DO;
                    DPRAM_Used_Payload.ISO_Rd   += TempMem;
                    DPRAM_Used_Payload.IRQ_Wr   += TempMemWr;
                    DOCounter.IRQ_Wr  += 1;

                end_case;

                DPRAM_Used_Payload.Payload_Read += TempMem;
                DPRAM_Used_Payload.Payload_Write += TempMemWr;

                if ud_DolType <> VARAN_DOL_IRQ then
                  DPRAM_Used.Total  += TempMem + TempMemWr + SIZE_PAYLOAD_FRAME_HEADER_DO;
                  DPRAM_Used_Payload.Payload_Header += SIZE_PAYLOAD_FRAME_HEADER_DO;
                else
                  DPRAM_Used.Total  += TempMem + TempMemWr + SIZE_PAYLOAD_IRQ_FRAME_HEADER_DO;
                  DPRAM_Used_Payload.Payload_Header += SIZE_PAYLOAD_IRQ_FRAME_HEADER_DO;
                end_if;

                DPRAM_Used_Payload.Total  += TempMem + TempMemWr;
                DOCounter.Total   += 1;

            VARAN_CMD_CONTROL_READ_WRITE,
            VARAN_CMD_MEMORY_READ_WRITE:// Read/Write DO -------------------------------------------------------------------------------------------------------------------------------
                // 1 Byte Control + n Byte (Load data read) + 0 to 3 Byte (compensate missalignment) x2
                TempMem := 1 + ud_ReadLength;

                TempMemWr := 1 + ud_WriteLength;

                // Increase for variable DO
                if ud_WritePayloadType = WR_PLD_TYPE_RW_ACCESS_CONFIGURABLE$UDINT then
                  TempMemWr += 16#13;
                elsif ud_WritePayloadType > WR_PLD_TYPE_STANDARD$UDINT then
                  TempMemWr += 16#0D;
                end_if;

                case ud_DolType of
                // **************************************************
                  VARAN_DOL_DA:
                    DPRAM_Used.DA_RdWr += TempMem + TempMemWr + SIZE_PAYLOAD_FRAME_HEADER_DO;
                    DPRAM_Used_Payload.DA_Rd += TempMem;
                    DPRAM_Used_Payload.DA_Wr += TempMemWr;
                    DOCounter.DA_RdWr  += 1;

                // **************************************************
                  VARAN_DOL_ISO:
                    DPRAM_Used.ISO_RdWr += TempMem + TempMemWr + SIZE_PAYLOAD_FRAME_HEADER_DO;
                    DPRAM_Used_Payload.ISO_Rd += TempMem;
                    DPRAM_Used_Payload.ISO_Wr += TempMemWr;

                    DOCounter.ISO_RdWr  += 1;

                // **************************************************
                  VARAN_DOL_ASY:
                    DPRAM_Used.ASY_RdWr += TempMem + TempMemWr + SIZE_PAYLOAD_FRAME_HEADER_DO;
                    DPRAM_Used_Payload.ASY_Rd += TempMem;
                    DPRAM_Used_Payload.ASY_Wr += TempMemWr;
                    DOCounter.ASY_RdWr  += 1;

                // **************************************************
                  VARAN_DOL_ADMIN:
                    DPRAM_Used.Admin_RdWr += TempMem + TempMemWr + SIZE_PAYLOAD_FRAME_HEADER_DO;
                    DPRAM_Used_Payload.Admin_Rd += TempMem;
                    DPRAM_Used_Payload.Admin_Wr += TempMemWr;
                    DOCounter.Admin_RdWr  += 1;

                // **************************************************
                  VARAN_DOL_IRQ:
                    DPRAM_Used.IRQ_RdWr += TempMem + TempMemWr + SIZE_PAYLOAD_IRQ_FRAME_HEADER_DO;
                    DPRAM_Used_Payload.IRQ_Rd += TempMem;
                    DPRAM_Used_Payload.IRQ_Wr += TempMemWr;
                    DOCounter.IRQ_RdWr  += 1;

                end_case;

                DPRAM_Used_Payload.Payload_Read += TempMem;
                DPRAM_Used_Payload.Payload_Write += TempMemWr;

                if ud_DolType <> VARAN_DOL_IRQ then
                  DPRAM_Used.Total  += TempMem + TempMemWr + SIZE_PAYLOAD_FRAME_HEADER_DO;
                  DPRAM_Used_Payload.Payload_Header += SIZE_PAYLOAD_FRAME_HEADER_DO;
                else
                  DPRAM_Used.Total  += TempMem + TempMemWr + SIZE_PAYLOAD_IRQ_FRAME_HEADER_DO;
                  DPRAM_Used_Payload.Payload_Header += SIZE_PAYLOAD_IRQ_FRAME_HEADER_DO;
                end_if;

                DPRAM_Used_Payload.Total += TempMem + TempMemWr;
                DOCounter.Total   += 1;

        end_case;
      else    // Standard DO Mem Calculation +++++++++++++++++++++++++++++++++++++++++++++++++++++++++++++++++++++++++++++++++++++++++++++++++++++++++++++++++++++++++++++++++++++++++

        case ud_Command of

            VARAN_CMD_CONTROL_READ,
            VARAN_CMD_MEMORY_READ:      // Read DO -------------------------------------------------------------------------------------------------------------------------------
                // 32 Byte (Header) + 6 Byte (1 Byte Cmd, 4 Byte Addr, 1 Byte Len) + 1 Byte (Response) + n Byte (Load data read) + 0 to 3 Byte (compensate missalignment)
                TempMem := 32 + 6 + 1 + ud_ReadLength;
                if (TempMem MOD 4) then
                  TempMem := TempMem + (4 - (TempMem MOD 4)); //increase memory, up to a value, which could be divided by 4
                end_if;

                case ud_DolType of
                // **************************************************
                  VARAN_DOL_DA:
                                DPRAM_Used.DA_Rd += TempMem;
                                DOCounter.DA_Rd  += 1;
                // **************************************************
                  VARAN_DOL_ISO:
                                DPRAM_Used.ISO_Rd += TempMem;
                                DOCounter.ISO_Rd  += 1;
                // **************************************************
                  VARAN_DOL_ASY:
                                DPRAM_Used.ASY_Rd += TempMem;
                                DOCounter.ASY_Rd  += 1;
                // **************************************************
                  VARAN_DOL_ADMIN:
                                DPRAM_Used.Admin_Rd += TempMem;
                                DOCounter.Admin_Rd  += 1;
                // **************************************************
                  VARAN_DOL_IRQ:
                                DPRAM_Used.IRQ_Rd += TempMem;
                                DOCounter.IRQ_Rd  += 1;
                end_case;

                DPRAM_Used.Total  += TempMem;
                DOCounter.Total   += 1;

            VARAN_CMD_CONTROL_WRITE,
            VARAN_CMD_MEMORY_WRITE:     // Write DO -------------------------------------------------------------------------------------------------------------------------------
                //32 Byte (Header) + 6 Byte (1 Byte Cmd, 4 Byte Addr, 1 Byte Len) + 1 Byte (Response) + n Byte (load data write) + 0 to 3 Byte (compensate missalignment)
                  TempMem := 32 + 6 + 1 + ud_WriteLength;
                  if (TempMem MOD 4) then
                    TempMem := TempMem + (4 - (TempMem MOD 4)); //increase memory, up to a value, which could be divided by 4
                  end_if;

                  case ud_DolType of
                  // **************************************************
                    VARAN_DOL_DA:
                                  DPRAM_Used.DA_Wr += TempMem;
                                  DOCounter.DA_Wr  += 1;
                  // **************************************************
                    VARAN_DOL_ISO:
                                  DPRAM_Used.ISO_Wr += TempMem;
                                  DOCounter.ISO_Wr  += 1;
                  // **************************************************
                    VARAN_DOL_ASY:
                                  DPRAM_Used.ASY_Wr += TempMem;
                                  DOCounter.ASY_Wr  += 1;
                  // **************************************************
                    VARAN_DOL_ADMIN:
                                  DPRAM_Used.Admin_Wr += TempMem;
                                  DOCounter.Admin_Wr  += 1;
                  // **************************************************
                    VARAN_DOL_IRQ:
                                  DPRAM_Used.IRQ_Wr += TempMem;
                                  DOCounter.IRQ_Wr  += 1;
                  end_case;

                  DPRAM_Used.Total  += TempMem;
                  DOCounter.Total   += 1;

            VARAN_CMD_CONTROL_READ_WRITE,
            VARAN_CMD_MEMORY_READ_WRITE:// Read/Write DO -------------------------------------------------------------------------------------------------------------------------------
                  //32 Byte (Header) + 11 Byte (1 Byte Cmd, 4 Byte RdAddr, 1 Byte RdLen, 4 Byte WrAddr, 1 Byte WrLen) + 1 Byte (Response) + n Byte (load data read) + n Byte (load data write) + 0 to 3 Byte (compensate missalignment)
                  TempMem := 32 + 11 + 1 + ud_ReadLength + ud_WriteLength;
                  if (TempMem MOD 4) then
                    TempMem := TempMem + (4 - (TempMem MOD 4)); //increase memory, up to a value, which could be divided by 4
                  end_if;

                  case ud_DolType of
                  // **************************************************
                    VARAN_DOL_DA:
                                  DPRAM_Used.DA_RdWr += TempMem;
                                  DOCounter.DA_RdWr  += 1;
                  // **************************************************
                    VARAN_DOL_ISO:
                                  DPRAM_Used.ISO_RdWr += TempMem;
                                  DOCounter.ISO_RdWr  += 1;
                  // **************************************************
                    VARAN_DOL_ASY:
                                  DPRAM_Used.ASY_RdWr += TempMem;
                                  DOCounter.ASY_RdWr  += 1;
                  // **************************************************
                    VARAN_DOL_ADMIN:
                                  DPRAM_Used.Admin_RdWr += TempMem;
                                  DOCounter.Admin_RdWr  += 1;
                  // **************************************************
                    VARAN_DOL_IRQ:
                                  DPRAM_Used.IRQ_RdWr += TempMem;
                                  DOCounter.IRQ_RdWr  += 1;
                  end_case;

                  DPRAM_Used.Total  += TempMem;
                  DOCounter.Total   += 1;

        end_case;

      end_if; // +++++++++++++++++++++++++++++++++++++++++++++++++++++++++++++++++++++++++++++++++++++++++++++++++++++++++++++++++++++++++++++++++++++++++++++++++++++++++++++++++++++++++++++++++

    end_if;
  else
    sd_retval := -100;	//Manager is off
  end_if;
END_FUNCTION

FUNCTION VaranManager::AddPayloadMoveDO
  VAR_INPUT
    p_ud_DoHandle 	: ^UDINT;
    ud_bDoRequired 	: UDINT;
    ud_DolType 	: UDINT;
    ud_Priority 	: UDINT;
    ud_PrescalerCounterThreshold 	: UDINT;
    ud_PrescalerCounterStartValue 	: UDINT;
    ud_hSourceReadDoHandle 	: UDINT;
    ud_ReadOffset 	: UDINT;
    ud_hDestinationWriteDoHandle 	: UDINT;
    ud_WriteOffset 	: UDINT;
    ud_MoveDataLength 	: UDINT;
  END_VAR
  VAR_OUTPUT
    sd_retval 	: DINT;
  END_VAR

#ifdef VM_DEBUG_PAYLOAD
  if b_PayloadSupport = false then
    // This method is not suppored without payload
    ((0)$^USINT)^ := 0;
  end_if;
#endif

  //look if we must execute Cyclic DOL list
  if ( ud_DolType = VARAN_DOL_ASY ) then
    s_CyHandles.b_ExecuteDOL := TRUE;			//set flag to execut Dol list
  end_if;

  sd_retval := MULTI_VARAN_iAddMoveDo(  phDoHandle                    := p_ud_DoHandle
                                      , bDoRequired                   := ud_bDoRequired
                                      , udDolType                     := ud_DolType
                                      , udPriority                    := ud_Priority
                                      , udPrescalerCounterThreshold   := ud_PrescalerCounterThreshold
                                      , udPrescalerCounterStartValue  := ud_PrescalerCounterStartValue
                                      , hSourceReadDoHandle           := ud_hSourceReadDoHandle
                                      , udReadOffset                  := ud_ReadOffset
                                      , hDestinationWriteDoHandle     := ud_hDestinationWriteDoHandle
                                      , udWriteOffset                 := ud_WriteOffset
                                      , udMoveDataLength              := ud_MoveDataLength);
  //look if an error occured
  if ( sd_retval <> VARANMANAGER_OK ) then
    s_ErrorVaranManager.f_AddRdDO := SetVaranDOError( sd_Error      := sd_retval
                                                    , b_manager_off := TRUE
                                                    , b_log         := TRUE
                                                    );
  else
    // Payload Move DO Mem Calculation
    if ( ud_DolType = VARAN_DOL_ASY ) then
      DPRAM_Used.ASY_Mov          += sizeof(LSL_VARANFRAMEPAYLOADMOVEHEADER);
      DPRAM_Used_Payload.ASY_Rd   += 1; // 1 Byte status
      DPRAM_Used_Payload.ASY_Wr   += sizeof(LSL_VARANFRAMEMOVEWRITEPAYLOAD);
      DOCounter.ASY_Mov           += 1;
    else
      DPRAM_Used.ISO_Mov          += sizeof(LSL_VARANFRAMEPAYLOADMOVEHEADER);
      DPRAM_Used_Payload.ISO_Rd   += 1; // 1 Byte status
      DPRAM_Used_Payload.ISO_Wr   += sizeof(LSL_VARANFRAMEMOVEWRITEPAYLOAD);
      DOCounter.ISO_Mov           += 1;
    end_if;

    DPRAM_Used.Total          += sizeof(LSL_VARANFRAMEPAYLOADMOVEHEADER) + 1 + sizeof(LSL_VARANFRAMEMOVEWRITEPAYLOAD);  // Header + Read Statusbyte + Write Payload
    DPRAM_Used_Payload.Total  += 1 + sizeof(LSL_VARANFRAMEMOVEWRITEPAYLOAD);  // Read Statusbyte + Write Payload
    DOCounter.Total           += 1;
  end_if;

END_FUNCTION

FUNCTION VaranManager::GetDataPointers
  VAR_INPUT
    ud_hDoHandle 	: UDINT;
    pp_ReadData 	: ^pVoid;
    pp_WriteData 	: ^pVoid;
  END_VAR
  VAR_OUTPUT
    sd_retval 	: DINT;
  END_VAR

#ifdef VM_DEBUG_PAYLOAD
  if b_PayloadSupport = false then
    // This method is not suppored without payload
    ((0)$^USINT)^ := 0;
  end_if;
#endif

  // if there is no VARAN Interface available, we would crash at the call
  if pMultiVaran = NIL then
    sd_retval := VARANMANAGER_DRIVER_NOT_EXISTS;
    return;
  end_if;

  sd_retval :=  MULTI_VARAN_iGetDataPointers( hDoHandle   := ud_hDoHandle
                                            , ppvReadData := pp_ReadData
                                            , ppvWriteData:= pp_WriteData);

END_FUNCTION

FUNCTION VaranManager::GetModuleHandle
  VAR_INPUT
    p_us_PositionInfo 	: ^USINT;
    p_ud_ModuleHandle 	: ^UDINT;
  END_VAR
  VAR_OUTPUT
    sd_retval 	: DINT;
  END_VAR

  // if there is no VARAN Interface available, we would crash at the call
  if pMultiVaran = NIL then
    sd_retval := VARANMANAGER_DRIVER_NOT_EXISTS;
    return;
  end_if;

  sd_retval := MULTI_VARAN_iGetNodeHandle(  udManagerNumber := VaranManagerNr
                                          , pszHardwarePath := p_us_PositionInfo
                                          , phNodeHandle    := p_ud_ModuleHandle);

END_FUNCTION

FUNCTION VaranManager::AddObjectCallback
	VAR_INPUT
		p_us_position_info 	: ^USINT;
		ud_action_ptr 	: UDINT;
		ud_thisp 	: UDINT;
		sd_required 	: DINT;
	END_VAR
	VAR_OUTPUT
		sd_retval 	: DINT;
	END_VAR
VAR
  ud_NodeHandle       :UDINT;
END_VAR

  if State = _NoVaranInterface then
    sd_retval := -100;
    return;
  end_if;
  //get right required flag
  if ( sd_required ) then
    sd_required := VARAN_DEVICE_REQUIRED;
  else
    sd_required := VARAN_DEVICE_DEFAULT;
  end_if;

    if b_PayloadSupport &
         _RTOSVersion >= VM_FULL_PAYLOAD_AVAILABLE  then
      sd_retval := MULTI_VARAN_iGetNodeHandle(  udManagerNumber := VaranManagerNr
                                              , pszHardwarePath := p_us_position_info
                                              , phNodeHandle    := #ud_NodeHandle);

      if sd_retval <> VARANMANAGER_OK then
        return;
      end_if;

      //call OS - function to set callback
      sd_retval := MULTI_VARAN_iSetApplicationCallback( hNodeHandle           := ud_NodeHandle
                                                      , pfApplicationCallback := ud_action_ptr$pvoid
                                                      , pvUserData            := ud_thisp$pvoid
                                                      , udRequired            := sd_required$UDINT);

    elsif pVaran then

      //call OS - function to set callback
      sd_retval := VARAN_iSetObjectCallback	( uiManager := VaranManagerNr
                                            , pucNode   := p_us_position_info
                                            , uiCallback:= ud_action_ptr
                                            , uiThis    := ud_thisp
                                            , uiRequired:= sd_required$UDINT
                                            );
    end_if;

  //look for an error
  if ( sd_retval <> VARANMANAGER_OK ) then
    s_ErrorVaranManager.f_SetObjectCallback := SetVaranDOError	( sd_Error 		:= sd_retval
                                                                , b_manager_off	:= TRUE
                                                                , b_log			:= TRUE
                                                                );
  end_if;

END_FUNCTION

FUNCTION VIRTUAL VaranManager::LogValue
	VAR_INPUT
		pString 	: ^CHAR;
		Value 	: UDINT;
		Value2 	: UDINT;(* := 16#FFFFFFFF *)
		Value3 	: UDINT;(* := 16#FFFFFFFF *)
	END_VAR
  VAR
    TempStr       : ARRAY [0..99] OF CHAR;
    TempStr2      : ARRAY [0..99] OF CHAR;
    TempStr3      : ARRAY [0..99] OF CHAR;
    TraceVal      : USINT;
    sz_name       : ARRAY [ 0..255 ] OF CHAR;
    TmpWithObjName: ARRAY [ 0..255 ] OF CHAR;
  END_VAR

  // number of values
  TraceVal := 1;

  _itoa(Value, #TempStr[0]);

  if pString <> NIL then
    _GetObjName( this, #sz_name[ 0 ] );
    _strcpy(dest:=#TmpWithObjName[0], src:="ObjectName ");
    _strcat(dest:=#TmpWithObjName[0], src:=#sz_name[0]);
    _strcat(dest:=#TmpWithObjName[0], src:=": ");
    _strcat(dest:=#TmpWithObjName[0], src:=pString);

    if Value2 <> 16#FFFFFFFF then
      _itoa(Value2, #TempStr2[0]);
      TraceVal += 1;
    end_if;

    if Value3 <> 16#FFFFFFFF then
      _itoa(Value3, #TempStr3[0]);
      TraceVal += 1;
    end_if;

    case TraceVal of
      1:MyTrace(pFormat:=#TmpWithObjName[0], pTxt0:=#TempStr[0], pTxt1:=NIL, pTxt2:=NIL);
      2:MyTrace(pFormat:=#TmpWithObjName[0], pTxt0:=#TempStr[0], pTxt1:=#TempStr2[0], pTxt2:=NIL);
      3:MyTrace(pFormat:=#TmpWithObjName[0], pTxt0:=#TempStr[0], pTxt1:=#TempStr2[0], pTxt2:=#TempStr3[0]);
    end_case;
  else
    MyTrace(pFormat:="<invalid string>", pTxt0:=NIL, pTxt1:=NIL, pTxt2:=NIL);
  end_if;

END_FUNCTION

FUNCTION VIRTUAL VaranManager::MyTrace
	VAR_INPUT
		pFormat 	: ^CHAR;
		pTxt0 	: ^CHAR;
		pTxt1 	: ^CHAR;
		pTxt2 	: ^CHAR;
	END_VAR
  VAR
    nLen      : UDINT;
    pChr      : ^CHAR;
    nTxt      : UDINT;
    nRpl      : UDINT;
    pTxt      : ^CHAR;
    pText     : ^CHAR;
    FormText  : ARRAY [0 .. 255] OF CHAR;
  END_VAR

  // this method is a workaround for the TRACE message limitation problem

  pText := #FormText[0];

  _memset(dest:=#FormText[0], usByte:=0, cntr:=256); // to keep the zero termination

  _strncpy(pText, pFormat, 250);
  nLen  := _strlen(pText);
  pChr  := pText;

  WHILE nLen DO
    IF pChr^ = '{' THEN         // works for the first 10 replacement texts (single digit numbers)
      nTxt  := (pChr+1)^ - '0';
      CASE nTxt OF
        0:  pTxt  := pTxt0;
        1:  pTxt  := pTxt1;
        2:  pTxt  := pTxt2;
      ELSE
        pTxt  := "INV";
      END_CASE;
      nRpl  := _strlen(pTxt);
      if nLen - 3 + nRpl > 250 then
        pTxt := "LEN";  // replace the replacement text with "LEN" to see that we're out of length for this string
        nRpl := 3;
      end_if;
      _memmove(pChr + nRpl, pChr + 3, nLen);
      _memcpy(pChr, pTxt, nRpl);
      pChr  += nRpl;  // next character to parse is after the replacement text
      nLen  -= 3;     // the remaining length of the format string is decremented by 3
      if nLen > 250 then  // catch overrun of nLen
        nLen := 0;
      end_if;
    ELSE
      pChr  += 1;
      nLen  -= 1;
    END_IF;
  END_WHILE;

  TRACE(#FormText[0]);
  if ( p_KernelLog ) then
    OS_KERNELLOG0(#FormText[0]);
  end_if;

END_FUNCTION

FUNCTION VaranManager::GetSPIDataFromID
	VAR_INPUT
		p_us_position_info 	: ^USINT;
		udListID 	: UDINT;
		pData 	: ^CHAR;
		udRequDataLength 	: UDINT;
		pIDHeader 	: ^t_s_SPIListHeader;
		udOffset 	: UDINT;(* := 16#00 *)
	END_VAR
	VAR_OUTPUT
		sd_retval 	: DINT;
	END_VAR

  VAR
    BaseListAddress : UDINT;
    a_data  : ARRAY[0..31] OF UDINT;
  END_VAR

  if p_us_position_info & pData & udRequDataLength > 0 then

    //check OS version
    if ( _RTOSVersion < VM_SPI_OS_VERSION ) then
      // access of SPI flash not possible
      sd_retval := -2;
      return;
    end_if;

    // check if list is available and get size and offset in SPI flash
    if ( SearchSPIList(p_us_position_info, udListID, #BaseListAddress) <> VARANMANAGER_OK ) then
      sd_retval := -3;
      return;
    end_if;

    //read header of list
    sd_retval := ReadSPIDataComfort(p_us_position_info := p_us_position_info,
                                    ud_offset := BaseListAddress,
                                    ud_length	:= sizeof(t_s_SPIListHeader),
                                    p_data	:= ( #a_data )$^USINT
                                    );

    _memcpy(ptr1:=pIDHeader, ptr2:=#a_data[0], cntr:=sizeof(t_s_SPIListHeader));

    //look for an error and check if length is > 0
    if ( sd_retval <> VARANMANAGER_OK ) | ( a_data[ 2 ] = 0 ) then
      sd_retval := -4;
      return;
    end_if;

    //read the whole serial number string
    sd_retval := ReadSPIDataComfort( p_us_position_info := p_us_position_info,
                                     ud_offset	:= BaseListAddress + sizeof(t_s_SPIListHeader) + udOffset,  //+12 ist List Header
                                     ud_length	:= udRequDataLength,
                                     p_data		:= pData
                                    );

    //look for an error
    if ( sd_retval <> VARANMANAGER_OK ) then
      sd_retval := -5;
      return;
    end_if;
  else
    // invalid parameters
    sd_retval := -1;
  end_if;

END_FUNCTION

FUNCTION GLOBAL VaranManager::RaiseManagerError
	VAR_INPUT
		udReason 	: UDINT;
	END_VAR

  State := udReason$t_e_VaranErrors;

  if b_PayloadSupport & _RTOSVersion >= VM_FULL_PAYLOAD_AVAILABLE  then
    MULTI_VARAN_iReportVaranError(diErrorNumber := udReason$DINT
                                , hErrorNode    := vmNodeHandle);

  elsif pVaran & (pVaran^.udVersion >= 16#00001104 ) then
    VARAN_iSetManagerError( VaranManagerNr, udReason );
  end_if;

END_FUNCTION
